(*
SPDX-FileCopyrightText: c 2026 Oleksandr Tiutyk <trofimich@gmail.com>
SPDX-License-Identifier: MIT
License: https://opensource.org/license/mit
*)

(*!
<summary>Checks that all three logger types contain an exception raised by the message formatter.</summary>
<description>
The runner task owns the fixtures. Each run clears its observations and uses the same instances. The file
logger remains idle in INITIAL without cyclic service.
</description>
*)

{attribute 'no_assign'}
{attribute 'no_explicit_call' := 'do not call this function block directly'}
FUNCTION_BLOCK LoggerFormatterFailureTest EXTENDS TOF_Testing.SingleCycleTest
VAR_STAT
	{attribute 'hide'}
	_ClassName : STRING := __POUNAME();
END_VAR
VAR
	_Queue : TOF_Loggers.QueuedLogger;
	_Backend : LoggerCaptureBackend;
	_EventLogger : TOF_Loggers.EventLogger(
		debugEventType := TC_EVENTS.OpenFrameworkLoggerEventClass.DebugEvent,
		informationEventType := TC_EVENTS.OpenFrameworkLoggerEventClass.InformationEvent,
		warningEventType := TC_EVENTS.OpenFrameworkLoggerEventClass.WarningEvent,
		errorEventType := TC_EVENTS.OpenFrameworkLoggerEventClass.ErrorEvent,
		criticalErrorEventType := TC_EVENTS.OpenFrameworkLoggerEventClass.CriticalErrorEvent
	);
	_FileLogger : TOF_Loggers.SimpleTextFileLogger(
		directoryPath := '',
		logFilePrefix := 'Log',
		maxRecordsPerFile := 1,
		directoryPathType := Tc2_System.E_OpenPath.PATH_GENERIC,
		timeout := T#2S,
		amsNetId := ''
	);
	_Formatter : ThrowingGetMessageException;
	_QueueConfigured : BOOL;
END_VAR

(*!
<summary>Checks that all three logger types contain an exception raised by the message formatter.</summary>
<description>
The runner task owns the fixtures. Each run clears its observations and uses the same instances. The file
logger remains idle in INITIAL without cyclic service.
</description>
*)
METHOD PROTECTED ExecuteTest
VAR
	formatCallsBefore : UDINT;
END_VAR
IF NOT _QueueConfigured THEN
	_QueueConfigured := _Queue.Configure(backend := _Backend);
END_IF

Assert.ThatBool(actual := _QueueConfigured, message := "Queue must bind to its capture backend").IsTrue();

IF NOT _QueueConfigured THEN
	RETURN;
END_IF

Assert.ThatBool(
	actual := _Queue.PendingMessageCount = 0,
	message := "Scenario must start with an empty queue"
).IsTrue();
formatCallsBefore := _Formatter.MessageReadCount;
Assert.ThatBool(
	actual := _Queue.TryLogException(exception := _Formatter, severity := TOF_Core.ERROR_SEVERITY.ERROR),
	message := "Queued logger must contain a throwing formatter"
).IsFalse();
Assert.ThatUDInt(
	actual := _Formatter.MessageReadCount,
	message := "Queued logger must reach the throwing formatter"
).ToBe(expected := formatCallsBefore + 1);

formatCallsBefore := _Formatter.MessageReadCount;
Assert.ThatBool(
	actual := _FileLogger.TryLogException(exception := _Formatter, severity := TOF_Core.ERROR_SEVERITY.ERROR),
	message := "File logger must contain a throwing formatter before admission"
).IsFalse();
Assert.ThatUDInt(
	actual := _Formatter.MessageReadCount,
	message := "File logger must reach the throwing formatter"
).ToBe(expected := formatCallsBefore + 1);

formatCallsBefore := _Formatter.MessageReadCount;
Assert.ThatBool(
	actual := _EventLogger.TryLogException(exception := _Formatter, severity := TOF_Core.ERROR_SEVERITY.ERROR),
	message := "Event logger must contain a throwing formatter before native send"
).IsFalse();
Assert.ThatUDInt(
	actual := _Formatter.MessageReadCount,
	message := "Event logger must reach the throwing formatter"
).ToBe(expected := formatCallsBefore + 1);

Assert.ThatBool(
	actual := _Queue.PendingMessageCount = 0,
	message := "Failed formatting must not enqueue a record"
).IsTrue();
Assert.ThatBool(actual := _FileLogger.Busy, message := "INITIAL must still report pending initialization").IsTrue();
Assert.ThatBool(
	actual := _FileLogger.State = TOF_Loggers.SIMPLE_TEXT_FILE_LOGGER_STATE.INITIAL,
	message := "A formatting refusal must leave the file logger in INITIAL"
).IsTrue();
END_METHOD

(*!
<summary>Clears capture observations and injected faults before each run.</summary>
*)
METHOD PROTECTED BeforeTest
_Backend.ResetCapture();
END_METHOD

//! <summary>Borrows the concrete class name for the instance lifetime. Callers must not modify it.</summary>
{attribute 'monitoring' := 'call'}
PROPERTY ClassName : REFERENCE TO STRING
GET
ClassName REF= _ClassName;
END_GET
END_PROPERTY

//! <summary>Borrows the compiler-initialized namespace. Callers must not modify it.</summary>
{attribute 'monitoring' := 'call'}
PROPERTY NamespaceName : REFERENCE TO STRING
GET
NamespaceName REF= CurrentNamespace.Name;
END_GET
END_PROPERTY

//! <summary>Reports the complete instance size in bytes, excluding separately allocated storage.</summary>
{attribute 'monitoring' := 'call'}
PROPERTY SelfSize : ULINT
GET
SelfSize := XSIZEOF(THIS^);
END_GET
END_PROPERTY

END_FUNCTION_BLOCK

(* stored: Version 1.1.0.1
   POU LoggerFormatterFailureTest: Id {a3d8f603-ec0f-4d15-abb1-16e174fc5993}, SpecialFunc None
   Method ExecuteTest: Id {78cdd936-e619-4f2a-a661-5b499fcce655}
   Method BeforeTest: Id {24106d99-2b4e-4ce0-a750-3174e2f234d3}
   Property ClassName: Id {8139d3c7-a498-4cc8-8a4d-1508d998b0d4}
   Get Get: Id {593da199-4dfa-455a-bf1d-3add02f853c0}
   Property NamespaceName: Id {0a088407-315d-4e9e-827c-9a2900ef2aab}
   Get Get: Id {6e98f80e-e9c9-49ab-8846-7552786dcdf7}
   Property SelfSize: Id {116881b8-20c2-409d-9b4f-e36b2eb833a2}
   Get Get: Id {8d173ba0-c490-4098-b155-1c760d8705c7} *)
